FUNCTION_BLOCK ResetLedControl (* Basic Function Block Type *)
  (* Standard: 61499-2 *)
  (* Version 0.0, 10/21/2026, macie, Schneider Electric, Template *)
  PACKAGE Main;
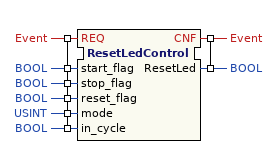
  EVENT_INPUT
    REQ WITH stop_flag, reset_flag, mode, in_cycle, start_flag; (* Normal Execution Request *)
  END_EVENT
  EVENT_OUTPUT
    CNF WITH ResetLed; (* Execution Confirmation *)
  END_EVENT
  VAR_INPUT
    start_flag : BOOL;
    stop_flag : BOOL; (* Input event qualifier *)
    reset_flag : BOOL;
    mode : USINT;
    in_cycle : BOOL;
  END_VAR
  VAR_OUTPUT
    ResetLed : BOOL; (* Output event qualifier *)
  END_VAR
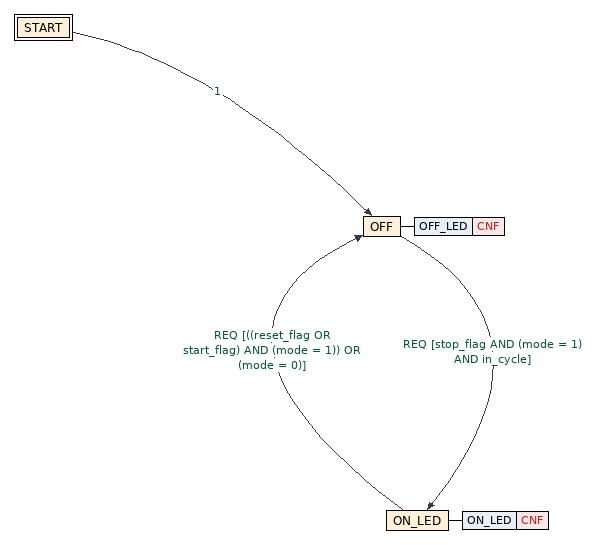
  EC_STATES
    START; (* Initial State *)
    OFF : OFF_LED -> CNF; (* Normal execution *)
    ON_LED : ON_LED -> CNF;
  END_STATES
  EC_TRANSITIONS
    START TO OFF := 1;
    OFF TO ON_LED := REQ [stop_flag AND (mode = 1) AND in_cycle];
    ON_LED TO OFF := REQ [((reset_flag OR start_flag) AND (mode = 1)) OR (mode = 0)];
  END_TRANSITIONS
  ALGORITHM ON_LED IN ST: (* Initialization algorithm *)
;
ResetLed := TRUE;
  END_ALGORITHM
  ALGORITHM OFF_LED IN ST: (* Normally executed algorithm *)
;
ResetLed := FALSE;
  END_ALGORITHM
END_FUNCTION_BLOCK
